// TIA Portal V21 export
Screen "R07_MoveV"  1024x768, Number=47, Template=Tpl
  ScreenLayer 
    Rectangle "P_CraneY" at 10,10 size 100x30
      VerticalMovementAnimation "VerticalMovementAnimation"
